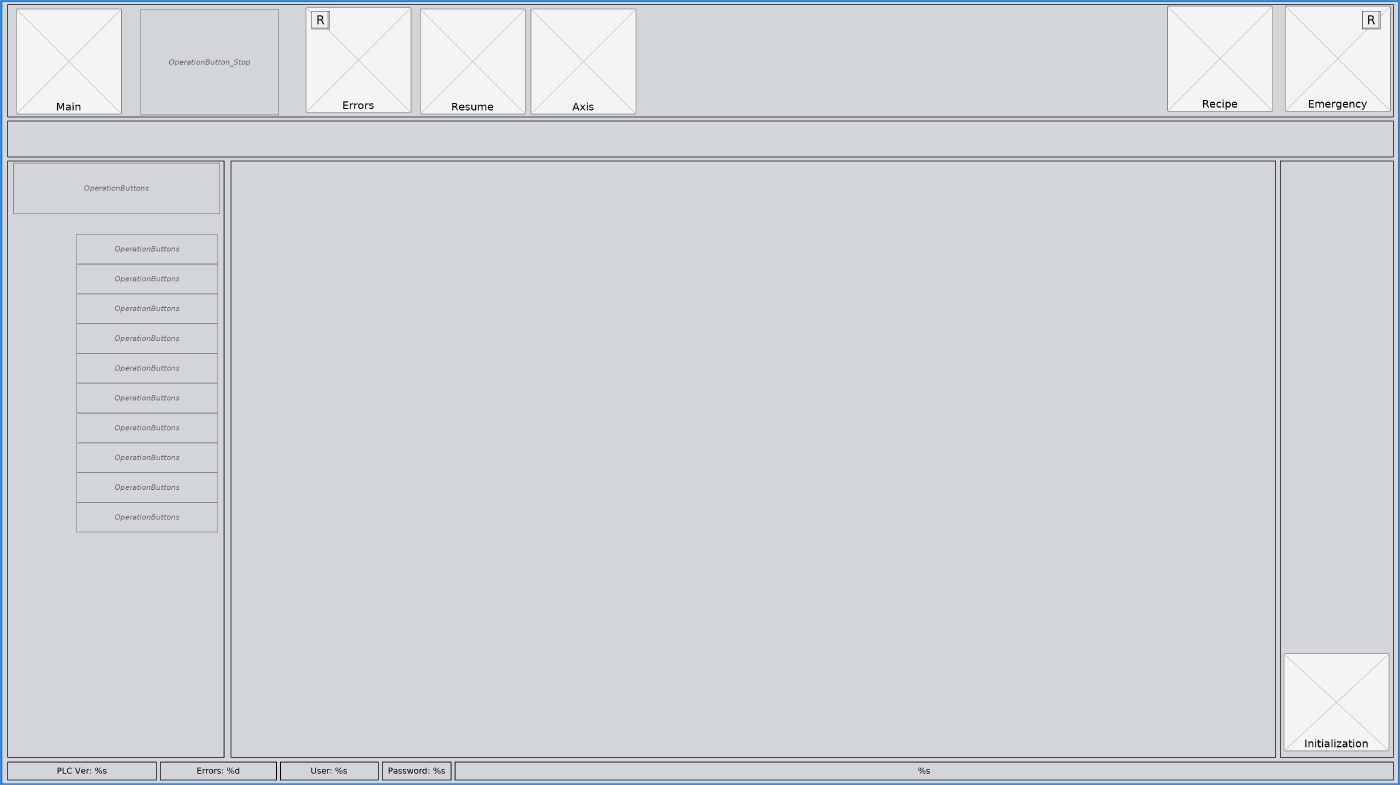
VISUALIZATION TEMP16_9_00  // 1924x1080
    Rectangle (0,0 1924x1080)
    Rectangle (385,1048 135x25), "User: %s", text variable: prg_User.actUser
    Rectangle (525,1048 95x25), "Password: %s", text variable: prg_User.Password
        OnMouseDown: write the text variable via Edit, min 1, max 999
    Rectangle (220,1048 160x25), "Errors: %d", text variable: Global_Persistent.Errors, colour toggle: Global_Persistent.Errors<>0
        OnMouseUp: execute { Global_Persistent.Errors:=(0); }
    Rectangle (10,1048 205x25), "PLC Ver: %s", text variable: ProgramVersion
    Rectangle (625,1048 1290x25), "%s", text variable: sDateTime
    Rectangle (10,6 1905x155)
    Rectangle (10,166 1905x50)
    Image (22,12 145x145), "Main", image: ImagePool.Main
        OnMouseClick: change screen: vis_MAIN
    Image (1766,8 145x145), "Emergency", image: ImagePool.EStop_OK2
        p84334746: GVL_Safety.sBitmap_ESButton
        OnMouseClick: change screen: ES_INT_OPER_16_9
    Image (420,10 145x145), "Errors", image: ImagePool.Error_No
        p84334746: s_Error_BitmapID
        OnMouseClick: change screen: ERRORS_OPER_16_9
    Image (577,12 145x145), "Resume", image: ImagePool.Resume3
        OnMouseClick: toggle ResumeAll
    Button (428,15 25x25), "R", pressed state: prg_Messages.ResetErrors
        toggle prg_Messages.ResetErrors
    Button (1872,15 25x25), "R"
    Rectangle (10,221 298x821)
    Rectangle (1759,221 156x821)
    Frame (18,224 284x70)
        shows OperationButtons(stOperation := stOpMain)
    Image (1764,899 145x134), "Initialization", image: ImagePool.illustration-project-icon
        OnMouseClick: change screen: INIT_OPER_16_9
    Rectangle (317,221 1436x821)
    Frame (193,13 190x145)
        shows OperationButton_Stop(stOperation := stOpMain)
    Image (729,12 145x145), "Axis", image: ImagePool.ervo-motor-beckhoff
        OnMouseClick: change screen: AXIS_OPER
    Image (1604,8 145x145), "Recipe", image: ImagePool.recipe icon
        OnMouseClick: change screen: Recipe_16_9
    Frame (105,322 194x41)
        shows OperationButtons(stOperation := stOper[E_ModeZone.eMain])
    Frame (105,363 194x41)
        shows OperationButtons(stOperation := stOper[E_ModeZone.eCIP])
    Frame (105,404 194x41)
        shows OperationButtons(stOperation := stOper[E_ModeZone.eTank1])
    Frame (105,445 194x41)
        shows OperationButtons(stOperation := stOper[E_ModeZone.eTank2])
    Frame (105,486 194x41)
        shows OperationButtons(stOperation := stOper[E_ModeZone.eTank3])
    Frame (105,527 194x41)
        shows OperationButtons(stOperation := stOper[E_ModeZone.eTank4])
    Frame (105,568 194x41)
        shows OperationButtons(stOperation := stOper[E_ModeZone.eProduction_Marinade])
    Frame (105,609 194x41)
        shows OperationButtons(stOperation := stOper[E_ModeZone.eProduction_Color])
    Frame (105,650 194x41)
        shows OperationButtons(stOperation := stOper[E_ModeZone.eTriBlender_Marinade])
    Frame (105,691 194x41)
        shows OperationButtons(stOperation := stOper[E_ModeZone.eTriBlender_Color])
END_VISUALIZATION

(* stored: Version 1.1.0.1, ProductVersion 3.1.4024.13
   Visu TEMP16_9_00: Id {5eaf349a-2f6b-4f8d-bd36-bc6832a62481} *)
